(* IEC 61131-3 sources: SafePLC-Gen-Evaluation/Evaluation Results/butane/run_01, 2 files *)

(* ---- io_declarations.st ---- *)
(* ==================================================  *)
(* PLC I/O Variable Declarations — CODESYS 3.5  *)
(* Generated by SafePLC-Gen Multimodal  *)
(* ==================================================  *)

VAR_GLOBAL
    (* --- Analog Inputs ---  *)
    TI_2909_Raw                  AT %IW0       : INT := 0;    (* TI-2909 — Temperature indicator, panel-mounted squ  *)
    TI_2917_Raw                  AT %IW2       : INT := 0;    (* TI-2917 — Temperature indicator with HH (high-high  *)
    TT_2909_Raw                  AT %IW4       : INT := 0;    (* TT-2909 — Temperature transmitter on inlet line up  *)
    TT_2911_Raw                  AT %IW6       : INT := 0;    (* TT-2911 — Temperature transmitter on outlet piping  *)
    TT_2917_Raw                  AT %IW8       : INT := 0;    (* TT-2917 — Temperature transmitter on utility/secon  *)
    XI_2901A_Raw                 AT %IW10      : INT := 0;    (* XI-2901A — Status indicator AVAILABLE for drive/MCC  *)
    XI_2901B_Raw                 AT %IW12      : INT := 0;    (* XI-2901B — Status indicator AVAILABLE for drive/MCC  *)
    (* --- Analog Outputs ---  *)
    HY_2903A_Out                 AT %QW0       : INT := 0;    (* HY-2903A — Hand relay/output converter for drive A,  *)
    HY_2903B_Out                 AT %QW2       : INT := 0;    (* HY-2903B — Hand relay/output converter for drive B,  *)
    (* --- Digital Inputs ---  *)
    ESD_3200                     AT %IX0.0     : BOOL := FALSE;    (* ESD-3200 — Emergency shutdown device/switch (ESD-32  *)
    HS_2901A                     AT %IX0.1     : BOOL := FALSE;    (* HS-2901A — Hand switch for drive A, panel-mounted s  *)
    HS_2901A1                    AT %IX0.2     : BOOL := FALSE;    (* HS-2901A1 — Hand switch LOCAL/REMOTE selector for dr  *)
    HS_2901A2                    AT %IX0.3     : BOOL := FALSE;    (* HS-2901A2 — Hand switch STOP/START for drive A, pane  *)
    HS_2901B                     AT %IX0.4     : BOOL := FALSE;    (* HS-2901B — Hand switch for drive B, panel-mounted s  *)
    HS_2901B1                    AT %IX0.5     : BOOL := FALSE;    (* HS-2901B1 — Hand switch LOCAL/REMOTE selector for dr  *)
    HS_2901B2                    AT %IX0.6     : BOOL := FALSE;    (* HS-2901B2 — Hand switch STOP/START for drive B, pane  *)
    HS_EMGSTOP_A_2901A           AT %IX0.7     : BOOL := FALSE;    (* HS-EMGSTOP-A-2901A — Hand switch EMERGENCY STOP (field-mounte  *)
    HS_EMGSTOP_B_2901B           AT %IX1.0     : BOOL := FALSE;    (* HS-EMGSTOP-B-2901B — Hand switch EMERGENCY STOP (field-mounte  *)
    HS_START_STOP_A_2901A        AT %IX1.1     : BOOL := FALSE;    (* HS-START-STOP-A-2901A — Hand switch START/STOP (field-mounted ci  *)
    HS_START_STOP_B_2901B        AT %IX1.2     : BOOL := FALSE;    (* HS-START-STOP-B-2901B — Hand switch START/STOP (field-mounted ci  *)
    PSD_2917                     AT %IX1.3     : BOOL := FALSE;    (* PSD-2917 — Pressure switch with shutdown function (  *)
    VSHH_2901A                   AT %IX1.4     : BOOL := FALSE;    (* VSHH-2901A — Vibration switch high-high on pump/compr  *)
    VSHH_2901B                   AT %IX1.5     : BOOL := FALSE;    (* VSHH-2901B — Vibration switch high-high on pump/compr  *)
    (* --- Digital Outputs ---  *)
    KV_2904                      AT %QX0.0     : BOOL := FALSE;    (* KV-2904 — Time-function valve or timer-operated va  *)
    XA_2901A                     AT %QX0.1     : BOOL := FALSE;    (* XA-2901A — Fault alarm indicator for drive A, panel  *)
    XA_2901B                     AT %QX0.2     : BOOL := FALSE;    (* XA-2901B — Fault alarm indicator for drive B, panel  *)
    XL_2901A                     AT %QX0.3     : BOOL := FALSE;    (* XL-2901A — Run status light/indicator RUNNING/STOP   *)
    XL_2901B                     AT %QX0.4     : BOOL := FALSE;    (* XL-2901B — Run status light/indicator RUNNING/STOP   *)
END_VAR

(* ---- generated_code.st ---- *)
(* Generated by SafePLC-Gen Multimodal — CODESYS 3.5 *)
(* IEC 61131-3 Structured Text *)
(* Date: 2026-04-25T12:02:41.596942 *)

PROGRAM PRG_Compressor_2901

VAR
    TI_2909_Raw             AT %IW0   : INT := 0;
    TI_2917_Raw             AT %IW2   : INT := 0;
    TT_2909_Raw             AT %IW4   : INT := 0;
    TT_2911_Raw             AT %IW6   : INT := 0;
    TT_2917_Raw             AT %IW8   : INT := 0;
    XI_2901A_Raw            AT %IW10  : INT := 0;
    XI_2901B_Raw            AT %IW12  : INT := 0;
    HY_2903A_Out            AT %QW0   : INT := 0;
    HY_2903B_Out            AT %QW2   : INT := 0;
    ESD_3200                AT %IX0.0 : BOOL := FALSE;
    HS_2901A                AT %IX0.1 : BOOL := FALSE;
    HS_2901A1               AT %IX0.2 : BOOL := FALSE;
    HS_2901A2               AT %IX0.3 : BOOL := FALSE;
    HS_2901B                AT %IX0.4 : BOOL := FALSE;
    HS_2901B1               AT %IX0.5 : BOOL := FALSE;
    HS_2901B2               AT %IX0.6 : BOOL := FALSE;
    HS_EMGSTOP_A_2901A      AT %IX0.7 : BOOL := FALSE;
    HS_EMGSTOP_B_2901B      AT %IX1.0 : BOOL := FALSE;
    HS_START_STOP_A_2901A   AT %IX1.1 : BOOL := FALSE;
    HS_START_STOP_B_2901B   AT %IX1.2 : BOOL := FALSE;
    PSD_2917                AT %IX1.3 : BOOL := FALSE;
    VSHH_2901A              AT %IX1.4 : BOOL := FALSE;
    VSHH_2901B              AT %IX1.5 : BOOL := FALSE;
    KV_2904                 AT %QX0.0 : BOOL := FALSE;
    XA_2901A                AT %QX0.1 : BOOL := FALSE;
    XA_2901B                AT %QX0.2 : BOOL := FALSE;
    XL_2901A                AT %QX0.3 : BOOL := FALSE;
    XL_2901B                AT %QX0.4 : BOOL := FALSE;
    ESTOP                   AT %IX2.0 : BOOL := FALSE;
    MANUAL_RESET            AT %IX2.1 : BOOL := FALSE;
END_VAR

VAR
    FirstScan               : BOOL := TRUE;

    TI_2909_Scaled          : REAL := 0.0;
    TT_2909_Scaled          : REAL := 0.0;
    TT_2911_Scaled          : REAL := 0.0;
    TT_2917_Scaled          : REAL := 0.0;
    TI_2917_Scaled          : REAL := 0.0;
    XI_2901A_Scaled         : REAL := 0.0;
    XI_2901B_Scaled         : REAL := 0.0;

    TI_2909_HH_SP           : REAL := 120.0;
    TI_2909_H_SP            : REAL := 110.0;
    TI_2909_L_SP            : REAL := 10.0;
    TI_2909_LL_SP           : REAL := 5.0;
    TI_2909_Deadband        : REAL := 2.0;
    TI_2909_HH_Latch        : BOOL := FALSE;
    TI_2909_LL_Latch        : BOOL := FALSE;
    TI_2909_HH              : BOOL := FALSE;
    TI_2909_H               : BOOL := FALSE;
    TI_2909_L               : BOOL := FALSE;
    TI_2909_LL              : BOOL := FALSE;
    TI_2909_HH_Ack          : BOOL := FALSE;
    TI_2909_LL_Ack          : BOOL := FALSE;

    TT_2909_HH_SP           : REAL := 120.0;
    TT_2909_H_SP            : REAL := 110.0;
    TT_2909_L_SP            : REAL := 10.0;
    TT_2909_LL_SP           : REAL := 5.0;
    TT_2909_Deadband        : REAL := 2.0;
    TT_2909_HH_Latch        : BOOL := FALSE;
    TT_2909_LL_Latch        : BOOL := FALSE;
    TT_2909_HH              : BOOL := FALSE;
    TT_2909_H               : BOOL := FALSE;
    TT_2909_L               : BOOL := FALSE;
    TT_2909_LL              : BOOL := FALSE;
    TT_2909_HH_Ack          : BOOL := FALSE;
    TT_2909_LL_Ack          : BOOL := FALSE;

    TT_2911_HH_SP           : REAL := 120.0;
    TT_2911_H_SP            : REAL := 110.0;
    TT_2911_L_SP            : REAL := 10.0;
    TT_2911_LL_SP           : REAL := 5.0;
    TT_2911_Deadband        : REAL := 2.0;
    TT_2911_HH_Latch        : BOOL := FALSE;
    TT_2911_LL_Latch        : BOOL := FALSE;
    TT_2911_HH              : BOOL := FALSE;
    TT_2911_H               : BOOL := FALSE;
    TT_2911_L               : BOOL := FALSE;
    TT_2911_LL              : BOOL := FALSE;
    TT_2911_HH_Ack          : BOOL := FALSE;
    TT_2911_LL_Ack          : BOOL := FALSE;

    TT_2917_HH_SP           : REAL := 130.0;
    TT_2917_H_SP            : REAL := 120.0;
    TT_2917_L_SP            : REAL := 10.0;
    TT_2917_LL_SP           : REAL := 5.0;
    TT_2917_Deadband        : REAL := 2.0;
    TT_2917_HH_Latch        : BOOL := FALSE;
    TT_2917_LL_Latch        : BOOL := FALSE;
    TT_2917_HH              : BOOL := FALSE;
    TT_2917_H               : BOOL := FALSE;
    TT_2917_L               : BOOL := FALSE;
    TT_2917_LL              : BOOL := FALSE;
    TT_2917_HH_Ack          : BOOL := FALSE;
    TT_2917_LL_Ack          : BOOL := FALSE;

    TI_2917_HH_SP           : REAL := 130.0;
    TI_2917_H_SP            : REAL := 120.0;
    TI_2917_L_SP            : REAL := 10.0;
    TI_2917_LL_SP           : REAL := 5.0;
    TI_2917_Deadband        : REAL := 2.0;
    TI_2917_HH_Latch        : BOOL := FALSE;
    TI_2917_LL_Latch        : BOOL := FALSE;
    TI_2917_HH              : BOOL := FALSE;
    TI_2917_H               : BOOL := FALSE;
    TI_2917_L               : BOOL := FALSE;
    TI_2917_LL              : BOOL := FALSE;
    TI_2917_HH_Ack          : BOOL := FALSE;
    TI_2917_LL_Ack          : BOOL := FALSE;

    XI_2901A_HH_SP          : REAL := 90.0;
    XI_2901A_H_SP           : REAL := 80.0;
    XI_2901A_L_SP           : REAL := 20.0;
    XI_2901A_LL_SP          : REAL := 10.0;
    XI_2901A_Deadband       : REAL := 2.0;
    XI_2901A_HH_Latch       : BOOL := FALSE;
    XI_2901A_LL_Latch       : BOOL := FALSE;
    XI_2901A_HH             : BOOL := FALSE;
    XI_2901A_H              : BOOL := FALSE;
    XI_2901A_L              : BOOL := FALSE;
    XI_2901A_LL             : BOOL := FALSE;
    XI_2901A_HH_Ack         : BOOL := FALSE;
    XI_2901A_LL_Ack         : BOOL := FALSE;

    XI_2901B_HH_SP          : REAL := 90.0;
    XI_2901B_H_SP           : REAL := 80.0;
    XI_2901B_L_SP           : REAL := 20.0;
    XI_2901B_LL_SP          : REAL := 10.0;
    XI_2901B_Deadband       : REAL := 2.0;
    XI_2901B_HH_Latch       : BOOL := FALSE;
    XI_2901B_LL_Latch       : BOOL := FALSE;
    XI_2901B_HH             : BOOL := FALSE;
    XI_2901B_H              : BOOL := FALSE;
    XI_2901B_L              : BOOL := FALSE;
    XI_2901B_LL             : BOOL := FALSE;
    XI_2901B_HH_Ack         : BOOL := FALSE;
    XI_2901B_LL_Ack         : BOOL := FALSE;

    LOOP_2917_TRIP          : BOOL := FALSE;
    LOOP_2901A_TRIP         : BOOL := FALSE;
    LOOP_2901B_TRIP         : BOOL := FALSE;
    VSHH_2901A_HH           : BOOL := FALSE;
    VSHH_2901A_LL           : BOOL := FALSE;
    VSHH_2901B_HH           : BOOL := FALSE;
    VSHH_2901B_LL           : BOOL := FALSE;
    SAFE_STATE              : BOOL := FALSE;

    MCC_A_Run               : BOOL := FALSE;
    MCC_B_Run               : BOOL := FALSE;
    MCC_A_Out               : BOOL := FALSE;
    MCC_B_Out               : BOOL := FALSE;

    Drive_A_SP              : REAL := 50.0;
    Drive_B_SP              : REAL := 50.0;
    Drive_A_Kp              : REAL := 1.0;
    Drive_A_Ki              : REAL := 0.1;
    Drive_B_Kp              : REAL := 1.0;
    Drive_B_Ki              : REAL := 0.1;
    Drive_A_Error           : REAL := 0.0;
    Drive_B_Error           : REAL := 0.0;
    Drive_A_Integral        : REAL := 0.0;
    Drive_B_Integral        : REAL := 0.0;
    Drive_A_Output          : REAL := 0.0;
    Drive_B_Output          : REAL := 0.0;

    StartDelay_A            : TON := (IN := FALSE, PT := T#3S);
    StartDelay_B            : TON := (IN := FALSE, PT := T#3S);

    RS_2901_Inlet_A_Upper   : BOOL := FALSE;
    RS_2901_Inlet_A_Lower   : BOOL := FALSE;
    RS_2901_Outlet_B_Upper  : BOOL := FALSE;
    RS_2901_Outlet_B_Lower  : BOOL := FALSE;
    BV_Inlet_A_Upper_1      : BOOL := FALSE;
    BV_Inlet_A_Upper_2      : BOOL := FALSE;
    BV_Inlet_A_Lower_1      : BOOL := FALSE;
    BV_Inlet_A_Lower_2      : BOOL := FALSE;
    BV_Outlet_B_Upper_1     : BOOL := FALSE;
    BV_Outlet_B_Upper_2     : BOOL := FALSE;
    BV_Outlet_B_Lower_1     : BOOL := FALSE;
    BV_Outlet_B_Lower_2     : BOOL := FALSE;
    CV_HY_2903A_1           : BOOL := FALSE;
    CV_HY_2903A_2           : BOOL := FALSE;
    CV_HY_2903B_1           : BOOL := FALSE;
    CV_HY_2903B_2           : BOOL := FALSE;
    CSO_Inlet_1             : BOOL := FALSE;
    CSO_Inlet_2             : BOOL := FALSE;
    FLV_Inlet               : BOOL := FALSE;
    BV_1IN_Drain            : BOOL := FALSE;
    Breather_A_8IN          : BOOL := FALSE;
    Breather_B_8IN          : BOOL := FALSE;
    NC_Valve_Outlet         : BOOL := FALSE;

    System_Alarm            : BOOL := FALSE;
END_VAR

IF FirstScan THEN
    LOOP_2917_TRIP          := TRUE;
    LOOP_2901A_TRIP         := TRUE;
    LOOP_2901B_TRIP         := TRUE;
    SAFE_STATE              := TRUE;
    MCC_A_Out               := FALSE;
    MCC_B_Out               := FALSE;
    MCC_A_Run               := FALSE;
    MCC_B_Run               := FALSE;
    HY_2903A_Out            := 6554;
    HY_2903B_Out            := 6554;
    KV_2904                 := FALSE;
    XL_2901A                := FALSE;
    XL_2901B                := FALSE;
    XA_2901A                := FALSE;
    XA_2901B                := FALSE;
    TI_2909_HH_Latch        := FALSE;
    TI_2909_LL_Latch        := FALSE;
    TT_2909_HH_Latch        := FALSE;
    TT_2909_LL_Latch        := FALSE;
    TT_2911_HH_Latch        := FALSE;
    TT_2911_LL_Latch        := FALSE;
    TT_2917_HH_Latch        := FALSE;
    TT_2917_LL_Latch        := FALSE;
    TI_2917_HH_Latch        := FALSE;
    TI_2917_LL_Latch        := FALSE;
    XI_2901A_HH_Latch       := FALSE;
    XI_2901A_LL_Latch       := FALSE;
    XI_2901B_HH_Latch       := FALSE;
    XI_2901B_LL_Latch       := FALSE;
    Drive_A_Integral        := 0.0;
    Drive_B_Integral        := 0.0;
    BV_1IN_Drain            := TRUE;
    StartDelay_A(IN := FALSE, PT := T#3S);
    StartDelay_B(IN := FALSE, PT := T#3S);
    FirstScan               := FALSE;
    RETURN;
END_IF;

TI_2909_Scaled  := ((INT_TO_REAL(TI_2909_Raw)  - 6554.0) / (32767.0 - 6554.0)) * 150.0;
TT_2909_Scaled  := ((INT_TO_REAL(TT_2909_Raw)  - 6554.0) / (32767.0 - 6554.0)) * 150.0;
TT_2911_Scaled  := ((INT_TO_REAL(TT_2911_Raw)  - 6554.0) / (32767.0 - 6554.0)) * 150.0;
TT_2917_Scaled  := ((INT_TO_REAL(TT_2917_Raw)  - 6554.0) / (32767.0 - 6554.0)) * 150.0;
TI_2917_Scaled  := ((INT_TO_REAL(TI_2917_Raw)  - 6554.0) / (32767.0 - 6554.0)) * 150.0;
XI_2901A_Scaled := ((INT_TO_REAL(XI_2901A_Raw) - 6554.0) / (32767.0 - 6554.0)) * 100.0;
XI_2901B_Scaled := ((INT_TO_REAL(XI_2901B_Raw) - 6554.0) / (32767.0 - 6554.0)) * 100.0;

IF TI_2909_Scaled >= TI_2909_HH_SP THEN
    TI_2909_HH_Latch := TRUE;
ELSIF TI_2909_Scaled <= (TI_2909_HH_SP - TI_2909_Deadband) AND TI_2909_HH_Ack THEN
    TI_2909_HH_Latch := FALSE;
END_IF;
TI_2909_HH := TI_2909_HH_Latch;
TI_2909_H  := TI_2909_Scaled >= TI_2909_H_SP;
TI_2909_L  := TI_2909_Scaled <= TI_2909_L_SP;
IF TI_2909_Scaled <= TI_2909_LL_SP THEN
    TI_2909_LL_Latch := TRUE;
ELSIF TI_2909_Scaled >= (TI_2909_LL_SP + TI_2909_Deadband) AND TI_2909_LL_Ack THEN
    TI_2909_LL_Latch := FALSE;
END_IF;
TI_2909_LL := TI_2909_LL_Latch;

IF TT_2909_Scaled >= TT_2909_HH_SP THEN
    TT_2909_HH_Latch := TRUE;
ELSIF TT_2909_Scaled <= (TT_2909_HH_SP - TT_2909_Deadband) AND TT_2909_HH_Ack THEN
    TT_2909_HH_Latch := FALSE;
END_IF;
TT_2909_HH := TT_2909_HH_Latch;
TT_2909_H  := TT_2909_Scaled >= TT_2909_H_SP;
TT_2909_L  := TT_2909_Scaled <= TT_2909_L_SP;
IF TT_2909_Scaled <= TT_2909_LL_SP THEN
    TT_2909_LL_Latch := TRUE;
ELSIF TT_2909_Scaled >= (TT_2909_LL_SP + TT_2909_Deadband) AND TT_2909_LL_Ack THEN
    TT_2909_LL_Latch := FALSE;
END_IF;
TT_2909_LL := TT_2909_LL_Latch;

IF TT_2911_Scaled >= TT_2911_HH_SP THEN
    TT_2911_HH_Latch := TRUE;
ELSIF TT_2911_Scaled <= (TT_2911_HH_SP - TT_2911_Deadband) AND TT_2911_HH_Ack THEN
    TT_2911_HH_Latch := FALSE;
END_IF;
TT_2911_HH := TT_2911_HH_Latch;
TT_2911_H  := TT_2911_Scaled >= TT_2911_H_SP;
TT_2911_L  := TT_2911_Scaled <= TT_2911_L_SP;
IF TT_2911_Scaled <= TT_2911_LL_SP THEN
    TT_2911_LL_Latch := TRUE;
ELSIF TT_2911_Scaled >= (TT_2911_LL_SP + TT_2911_Deadband) AND TT_2911_LL_Ack THEN
    TT_2911_LL_Latch := FALSE;
END_IF;
TT_2911_LL := TT_2911_LL_Latch;

IF TT_2917_Scaled >= TT_2917_HH_SP THEN
    TT_2917_HH_Latch := TRUE;
ELSIF TT_2917_Scaled <= (TT_2917_HH_SP - TT_2917_Deadband) AND TT_2917_HH_Ack THEN
    TT_2917_HH_Latch := FALSE;
END_IF;
TT_2917_HH := TT_2917_HH_Latch;
TT_2917_H  := TT_2917_Scaled >= TT_2917_H_SP;
TT_2917_L  := TT_2917_Scaled <= TT_2917_L_SP;
IF TT_2917_Scaled <= TT_2917_LL_SP THEN
    TT_2917_LL_Latch := TRUE;
ELSIF TT_2917_Scaled >= (TT_2917_LL_SP + TT_2917_Deadband) AND TT_2917_LL_Ack THEN
    TT_2917_LL_Latch := FALSE;
END_IF;
TT_2917_LL := TT_2917_LL_Latch;

IF TI_2917_Scaled >= TI_2917_HH_SP THEN
    TI_2917_HH_Latch := TRUE;
ELSIF TI_2917_Scaled <= (TI_2917_HH_SP - TI_2917_Deadband) AND TI_2917_HH_Ack THEN
    TI_2917_HH_Latch := FALSE;
END_IF;
TI_2917_HH := TI_2917_HH_Latch;
TI_2917_H  := TI_2917_Scaled >= TI_2917_H_SP;
TI_2917_L  := TI_2917_Scaled <= TI_2917_L_SP;
IF TI_2917_Scaled <= TI_2917_LL_SP THEN
    TI_2917_LL_Latch := TRUE;
ELSIF TI_2917_Scaled >= (TI_2917_LL_SP + TI_2917_Deadband) AND TI_2917_LL_Ack THEN
    TI_2917_LL_Latch := FALSE;
END_IF;
TI_2917_LL := TI_2917_LL_Latch;

IF XI_2901A_Scaled >= XI_2901A_HH_SP THEN
    XI_2901A_HH_Latch := TRUE;
ELSIF XI_2901A_Scaled <= (XI_2901A_HH_SP - XI_2901A_Deadband) AND XI_2901A_HH_Ack THEN
    XI_2901A_HH_Latch := FALSE;
END_IF;
XI_2901A_HH := XI_2901A_HH_Latch;
XI_2901A_H  := XI_2901A_Scaled >= XI_2901A_H_SP;
XI_2901A_L  := XI_2901A_Scaled <= XI_2901A_L_SP;
IF XI_2901A_Scaled <= XI_2901A_LL_SP THEN
    XI_2901A_LL_Latch := TRUE;
ELSIF XI_2901A_Scaled >= (XI_2901A_LL_SP + XI_2901A_Deadband) AND XI_2901A_LL_Ack THEN
    XI_2901A_LL_Latch := FALSE;
END_IF;
XI_2901A_LL := XI_2901A_LL_Latch;

IF XI_2901B_Scaled >= XI_2901B_HH_SP THEN
    XI_2901B_HH_Latch := TRUE;
ELSIF XI_2901B_Scaled <= (XI_2901B_HH_SP - XI_2901B_Deadband) AND XI_2901B_HH_Ack THEN
    XI_2901B_HH_Latch := FALSE;
END_IF;
XI_2901B_HH := XI_2901B_HH_Latch;
XI_2901B_H  := XI_2901B_Scaled >= XI_2901B_H_SP;
XI_2901B_L  := XI_2901B_Scaled <= XI_2901B_L_SP;
IF XI_2901B_Scaled <= XI_2901B_LL_SP THEN
    XI_2901B_LL_Latch := TRUE;
ELSIF XI_2901B_Scaled >= (XI_2901B_LL_SP + XI_2901B_Deadband) AND XI_2901B_LL_Ack THEN
    XI_2901B_LL_Latch := FALSE;
END_IF;
XI_2901B_LL := XI_2901B_LL_Latch;

VSHH_2901A_HH := VSHH_2901A;
VSHH_2901A_LL := FALSE;
VSHH_2901B_HH := VSHH_2901B;
VSHH_2901B_LL := FALSE;

IF TT_2917_HH OR TT_2917_LL OR TI_2917_HH OR TI_2917_LL OR PSD_2917 THEN
    LOOP_2917_TRIP := TRUE;
ELSIF LOOP_2917_TRIP AND MANUAL_RESET
      AND NOT TT_2917_HH AND NOT TT_2917_LL
      AND NOT TI_2917_HH AND NOT TI_2917_LL
      AND NOT PSD_2917 THEN
    LOOP_2917_TRIP := FALSE;
END_IF;

IF VSHH_2901A_HH OR VSHH_2901A_LL THEN
    LOOP_2901A_TRIP := TRUE;
ELSIF LOOP_2901A_TRIP AND MANUAL_RESET
      AND NOT VSHH_2901A_HH AND NOT VSHH_2901A_LL THEN
    LOOP_2901A_TRIP := FALSE;
END_IF;

IF VSHH_2901B_HH OR VSHH_2901B_LL THEN
    LOOP_2901B_TRIP := TRUE;
ELSIF LOOP_2901B_TRIP AND MANUAL_RESET
      AND NOT VSHH_2901B_HH AND NOT VSHH_2901B_LL THEN
    LOOP_2901B_TRIP := FALSE;
END_IF;

SAFE_STATE := ESTOP OR ESD_3200
              OR HS_EMGSTOP_A_2901A OR HS_EMGSTOP_B_2901B
              OR LOOP_2917_TRIP OR LOOP_2901A_TRIP OR LOOP_2901B_TRIP;

StartDelay_A(IN := MCC_A_Run AND NOT SAFE_STATE, PT := T#3S);
StartDelay_B(IN := MCC_B_Run AND NOT SAFE_STATE, PT := T#3S);

IF NOT SAFE_STATE THEN
    IF HS_2901A1 THEN
        IF HS_START_STOP_A_2901A THEN
            MCC_A_Run := TRUE;
        ELSIF NOT HS_2901A THEN
            MCC_A_Run := FALSE;
        END_IF;
    ELSE
        MCC_A_Run := HS_2901A2;
    END_IF;

    MCC_A_Out := StartDelay_A.Q;

    IF MCC_A_Out THEN
        Drive_A_Error    := Drive_A_SP - XI_2901A_Scaled;
        Drive_A_Integral := Drive_A_Integral + (Drive_A_Ki * Drive_A_Error);
        IF Drive_A_Integral > 100.0 THEN
            Drive_A_Integral := 100.0;
        ELSIF Drive_A_Integral < 0.0 THEN
            Drive_A_Integral := 0.0;
        END_IF;
        Drive_A_Output := (Drive_A_Kp * Drive_A_Error) + Drive_A_Integral;
        IF Drive_A_Output > 100.0 THEN
            Drive_A_Output := 100.0;
        ELSIF Drive_A_Output < 0.0 THEN
            Drive_A_Output := 0.0;
        END_IF;
        HY_2903A_Out := REAL_TO_INT(6554.0 + (Drive_A_Output / 100.0) * (32767.0 - 6554.0));
    ELSE
        HY_2903A_Out     := 6554;
        Drive_A_Integral := 0.0;
    END_IF;

    IF HS_2901B1 THEN
        IF HS_START_STOP_B_2901B THEN
            MCC_B_Run := TRUE;
        ELSIF NOT HS_2901B THEN
            MCC_B_Run := FALSE;
        END_IF;
    ELSE
        MCC_B_Run := HS_2901B2;
    END_IF;

    MCC_B_Out := StartDelay_B.Q;

    IF MCC_B_Out THEN
        Drive_B_Error    := Drive_B_SP - XI_2901B_Scaled;
        Drive_B_Integral := Drive_B_Integral + (Drive_B_Ki * Drive_B_Error);
        IF Drive_B_Integral > 100.0 THEN
            Drive_B_Integral := 100.0;
        ELSIF Drive_B_Integral < 0.0 THEN
            Drive_B_Integral := 0.0;
        END_IF;
        Drive_B_Output := (Drive_B_Kp * Drive_B_Error) + Drive_B_Integral;
        IF Drive_B_Output > 100.0 THEN
            Drive_B_Output := 100.0;
        ELSIF Drive_B_Output < 0.0 THEN
            Drive_B_Output := 0.0;
        END_IF;
        HY_2903B_Out := REAL_TO_INT(6554.0 + (Drive_B_Output / 100.0) * (32767.0 - 6554.0));
    ELSE
        HY_2903B_Out     := 6554;
        Drive_B_Integral := 0.0;
    END_IF;

    KV_2904                := MCC_A_Out OR MCC_B_Out;
    RS_2901_Inlet_A_Upper  := MCC_A_Out;
    RS_2901_Inlet_A_Lower  := MCC_A_Out;
    RS_2901_Outlet_B_Upper := MCC_B_Out;
    RS_2901_Outlet_B_Lower := MCC_B_Out;
    BV_Inlet_A_Upper_1     := MCC_A_Out;
    BV_Inlet_A_Upper_2     := MCC_A_Out;
    BV_Inlet_A_Lower_1     := MCC_A_Out;
    BV_Inlet_A_Lower_2     := MCC_A_Out;
    BV_Outlet_B_Upper_1    := MCC_B_Out;
    BV_Outlet_B_Upper_2    := MCC_B_Out;
    BV_Outlet_B_Lower_1    := MCC_B_Out;
    BV_Outlet_B_Lower_2    := MCC_B_Out;
    CV_HY_2903A_1          := MCC_A_Out;
    CV_HY_2903A_2          := MCC_A_Out;
    CV_HY_2903B_1          := MCC_B_Out;
    CV_HY_2903B_2          := MCC_B_Out;
    CSO_Inlet_1            := MCC_A_Out OR MCC_B_Out;
    CSO_Inlet_2            := MCC_A_Out OR MCC_B_Out;
    FLV_Inlet              := MCC_A_Out OR MCC_B_Out;
    BV_1IN_Drain           := NOT (MCC_A_Out OR MCC_B_Out);
    Breather_A_8IN         := MCC_A_Out;
    Breather_B_8IN         := MCC_B_Out;
    NC_Valve_Outlet        := MCC_A_Out OR MCC_B_Out;
    XL_2901A               := MCC_A_Out;
    XL_2901B               := MCC_B_Out;
    XA_2901A               := LOOP_2901A_TRIP OR XI_2901A_HH;
    XA_2901B               := LOOP_2901B_TRIP OR XI_2901B_HH;
ELSE
    MCC_A_Out              := FALSE;
    MCC_B_Out              := FALSE;
    MCC_A_Run              := FALSE;
    MCC_B_Run              := FALSE;
    HY_2903A_Out           := 6554;
    HY_2903B_Out           := 6554;
    KV_2904                := FALSE;
    XL_2901A               := FALSE;
    XL_2901B               := FALSE;
    XA_2901A               := TRUE;
    XA_2901B               := TRUE;
    Drive_A_Integral       := 0.0;
    Drive_B_Integral       := 0.0;
    RS_2901_Inlet_A_Upper  := FALSE;
    RS_2901_Inlet_A_Lower  := FALSE;
    RS_2901_Outlet_B_Upper := FALSE;
    RS_2901_Outlet_B_Lower := FALSE;
    BV_Inlet_A_Upper_1     := FALSE;
    BV_Inlet_A_Upper_2     := FALSE;
    BV_Inlet_A_Lower_1     := FALSE;
    BV_Inlet_A_Lower_2     := FALSE;
    BV_Outlet_B_Upper_1    := FALSE;
    BV_Outlet_B_Upper_2    := FALSE;
    BV_Outlet_B_Lower_1    := FALSE;
    BV_Outlet_B_Lower_2    := FALSE;
    CV_HY_2903A_1          := FALSE;
    CV_HY_2903A_2          := FALSE;
    CV_HY_2903B_1          := FALSE;
    CV_HY_2903B_2          := FALSE;
    CSO_Inlet_1            := FALSE;
    CSO_Inlet_2            := FALSE;
    FLV_Inlet              := FALSE;
    BV_1IN_Drain           := TRUE;
    Breather_A_8IN         := FALSE;
    Breather_B_8IN         := FALSE;
    NC_Valve_Outlet        := FALSE;
END_IF;

System_Alarm :=
    TI_2909_HH_Latch  OR TI_2909_LL_Latch  OR TI_2909_H  OR TI_2909_L  OR
    TT_2909_HH_Latch  OR TT_2909_LL_Latch  OR TT_2909_H  OR TT_2909_L  OR
    TT_2911_HH_Latch  OR TT_2911_LL_Latch  OR TT_2911_H  OR TT_2911_L  OR
    TT_2917_HH_Latch  OR TT_2917_LL_Latch  OR TT_2917_H  OR TT_2917_L  OR
    TI_2917_HH_Latch  OR TI_2917_LL_Latch  OR TI_2917_H  OR TI_2917_L  OR
    XI_2901A_HH_Latch OR XI_2901A_LL_Latch OR XI_2901A_H OR XI_2901A_L OR
    XI_2901B_HH_Latch OR XI_2901B_LL_Latch OR XI_2901B_H OR XI_2901B_L OR
    LOOP_2917_TRIP OR LOOP_2901A_TRIP OR LOOP_2901B_TRIP OR SAFE_STATE;

END_PROGRAM
